(* IEC 61131-3 sources: codesys-framework/txt/application/ToDo/Utils, 8 files *)

(* ---- E_ScaleMethod.dut.st ---- *)
TYPE E_ScaleMethod :
(
	InterPolationZero_whenOutLimits := 0,
	InterPolationLimitValue_whenOutLimits := 1,
	ExtraPolation := 2
);
END_TYPE

(* ---- E_TaskStatus.dut.st ---- *)
{attribute 'qualified_only'}
{attribute 'strict'}
TYPE E_TaskStatus :
(
	NotStarted := 0,		// Task has not yet began (default value)
	Start,					// Task start external request
	Busy,					// Task is busy
	Successful,				// Task ended successful
	Failed,					// Task ended failure
	Tolerated,				// Task ended failure, but failure is tolerated
	Error,					// Task experiences error
	Interrupted,			// Task was interrupted
	Skipped,				// Task was skipped
	Timeout					// Task timed out
);
END_TYPE

(* ---- F_GetEngUnit.pou.st ---- *)
FUNCTION F_GetEngUnit : STRING (20)
VAR_INPUT
	eEngUnit : E_EngineeringUnits;
END_VAR
VAR
	sEngUnitString : STRING(20);
END_VAR

// --- BEGIN IMPLEMENTATION ---

//Add EngineeringUnitString
CASE (eEngUnit) OF
	E_EngineeringUnits.Volt : sEngUnitString := 'V';
	E_EngineeringUnits.gram : sEngUnitString := 'gram';
	E_EngineeringUnits.bar : sEngUnitString := 'bar';
	E_EngineeringUnits.degree : sEngUnitString := '°';
	E_EngineeringUnits.cubicmeters : sEngUnitString := 'm³';
	E_EngineeringUnits.milimeters : sEngUnitString := 'mm';
	ELSE sEngUnitString := '';
END_CASE

F_GetEngUnit := sEngUnitString;

(* ---- F_Scale.pou.st ---- *)
FUNCTION F_Scale : REAL
VAR_INPUT
	rInputScaleValue : REAL;
	rInputScaleValueMinLevel : REAL;
	rInputScaleValueMaxLevel : REAL;
	rOutputScaleValueMinLevel : REAL;
	rOutputScaleValueMaxLevel : REAL;
	eScaleMethod : E_ScaleMethod;
END_VAR
VAR_OUTPUT
	xInputScaleValueBelowMinLevel : BOOL;
	xInputScaleValueAboveMaxLevel : BOOL;
	xInputScaleMinMaxDivisionByZero : BOOL;
END_VAR
VAR
	_rPercentValue : REAL;
END_VAR

// --- BEGIN IMPLEMENTATION ---

// Scale the <rInputScale_Value> between <rOutputScale_Value_MinLevel> and <rOutputScale_Value_MaxLevel>
// -- <rOutputScale_Value_MinLevel> ~ <rInputScale_Value_MinLevel>
// -- <rOutputScale_Value_MaxLevel> ~ <rInputScale_Value_MaxLevel>

// Check boundaries <nInputScale_Value>
xInputScaleValueBelowMinLevel := rInputScaleValue < rInputScaleValueMinLevel;
xInputScaleValueAboveMaxLevel := rInputScaleValue > rInputScaleValueMaxLevel;
xInputScaleMinMaxDivisionByZero := (rInputScaleValueMaxLevel - rInputScaleValueMinLevel) = 0;

// If error
IF eScaleMethod = E_ScaleMethod.InterPolationLimitValue_whenOutLimits AND (xInputScaleValueBelowMinLevel OR xInputScaleValueAboveMaxLevel) THEN

	IF xInputScaleValueBelowMinLevel THEN
		F_Scale := rOutputScaleValueMinLevel;

	ELSIF xInputScaleValueAboveMaxLevel THEN
		F_Scale := rOutputScaleValueMaxLevel;

	END_IF

ELSIF (eScaleMethod = E_ScaleMethod.InterPolationZero_whenOutLimits AND (xInputScaleValueBelowMinLevel OR xInputScaleValueAboveMaxLevel)) OR xInputScaleMinMaxDivisionByZero THEN
	F_Scale := 0.0;
ELSE
	_rPercentValue := (rInputScaleValue - rInputScaleValueMinLevel) / (rInputScaleValueMaxLevel - rInputScaleValueMinLevel);
	F_Scale := rOutputScaleValueMinLevel + ((rOutputScaleValueMaxLevel - rOutputScaleValueMinLevel) * _rPercentValue);
END_IF

(* ---- Round.pou.st ---- *)
FUNCTION Round : LREAL
VAR_INPUT
	lrValue 		: LREAL;
 	iDecimalPlaces 	: INT;
END_VAR
VAR
	_lrOutput 		: LREAL;
	_lrRightPart 	: LREAL;
  	_lrLeftPart 	: LREAL;
END_VAR

// --- BEGIN IMPLEMENTATION ---

_lrOutput := lrValue * EXPT(10, iDecimalPlaces);
_lrRightPart := DINT_TO_LREAL(TRUNC(_lrOutput));
_lrLeftPart := _lrOutput - _lrRightPart;

_lrOutput := _lrRightPart;

IF _lrLeftPart >= 0.5 THEN
  _lrOutput := _lrRightPart + 1;
END_IF

_lrOutput := _lrOutput / EXPT(10, iDecimalPlaces);

Round := _lrOutput;

(* ---- FB_CycleInfo.pou.st ---- *)
FUNCTION_BLOCK FB_CycleInfo
VAR_INPUT
	udiCycleStartEventID : UDINT;
END_VAR
VAR_OUTPUT
	rCycleTime_msec : REAL;
	udiCycleFirstStartCounter : UDINT;
END_VAR
VAR_IN_OUT
	xFirstCycleDone : BOOL;
	xResetFirstCycle : BOOL;
END_VAR
VAR
	_xFirstCycleNew : BOOL;
END_VAR

// --- BEGIN IMPLEMENTATION ---

IF xFirstCycleDone AND xResetFirstCycle THEN
	xResetFirstCycle := FALSE;
	_xFirstCycleNew := TRUE;
END_IF

IF NOT xFirstCycleDone AND xResetFirstCycle THEN
	xFirstCycleDone := TRUE;
END_IF

IF NOT xFirstCycleDone OR _xFirstCycleNew THEN
	xFirstCycleDone := FALSE;
	_xFirstCycleNew := FALSE;
	F_Event_InsertMessage (
		eSubMachine := 0,
		w := 1,
		iComponentID := 0,
		udiEventID := udiCycleStartEventID,
		eEventLevel := E_EventLevels.EventIsInformational);
	udiCycleFirstStartCounter := udiCycleFirstStartCounter + 1;
END_IF

(* ---- FB_GetIpAddress.pou.st ---- *)
FUNCTION_BLOCK FB_GetIpAddress
VAR_INPUT
END_VAR
VAR_OUTPUT
END_VAR
VAR
	_fbL_IPAP_ParameterRead		: L_IPAP_ParameterRead;

	_xRead 						: BOOL;
	_udiIp						: UDINT;
	_b1, _b2, _b3, _b4 			: BYTE;
	_sIp 						: STRING;
END_VAR

// --- BEGIN IMPLEMENTATION ---

_fbL_IPAP_ParameterRead(
	xExecute		:= _xRead ,
	xAbort			:= ,
	wIndex			:= 9298,
	bySubIndex		:= 1,
	udiTimeOut		:= 1000,
	pDataBuffer		:= ADR(_udiIp),
	udiBufferSize	:= SIZEOF(_udiIp),
	xDone			=> ,
	xBusy			=> ,
	xAborted		=> ,
	xError			=> ,
	eErrorId		=> ,
	udiDataRead		=> ,
	eDataType		=>
);

IF _xRead AND _fbL_IPAP_ParameterRead.xDone THEN
	 _xRead := FALSE;
END_IF

_b1 := TO_BYTE(SHR(_udiIp, 24));
_b2 := TO_BYTE(SHR(_udiIp, 16));
_b3 := TO_BYTE(SHR(_udiIp, 8));
_b4 := TO_BYTE(_udiIp);

_sIp := '';
_sIp := CONCAT(str1 := _sIp, str2 := TO_STRING(_b4));
_sIp := CONCAT(str1 := _sIp, str2 := '.');
_sIp := CONCAT(str1 := _sIp, str2 := TO_STRING(_b3));
_sIp := CONCAT(str1 := _sIp, str2 := '.');
_sIp := CONCAT(str1 := _sIp, str2 := TO_STRING(_b2));
_sIp := CONCAT(str1 := _sIp, str2 := '.');
_sIp := CONCAT(str1 := _sIp, str2 := TO_STRING(_b1));

(* ---- FB_Timer.pou.st ---- *)
FUNCTION_BLOCK FB_Timer
VAR_INPUT
END_VAR
VAR_OUTPUT
END_VAR
VAR
	_xOn 			: BOOL;
	_rtrigOn 		: R_TRIG;
	_ftrigOn 		: F_TRIG;

	_tStart 		: TIME;
	_tEnd 			: TIME;
	_tDelta 		: TIME;
	_tPrevious 		: TIME;
	_tTotal 		: TIME;
END_VAR

// --- BEGIN IMPLEMENTATION ---

_rtrigOn(CLK := _xOn);
_ftrigOn(CLK := _xOn);

IF _rtrigOn.Q THEN
	_tStart := TO_TIME(SysTimeGetMs());
END_IF

IF _ftrigOn.Q THEN
	_tPrevious := _tPrevious + _tDelta;
	_tDelta := T#0MS;
END_IF

IF _xOn THEN
	_tEnd := TO_TIME(SysTimeGetMs());
	_tDelta := _tEnd - _tStart;
END_IF

_tTotal := _tPrevious + _tDelta;
